PROGRAM prg_Call_Recipe_Slow
VAR
	i							: INT;
	bFirstScan					: BOOL:= TRUE;
	ton_RecipeReady				: TON;
	
	
	eRecipeName: E_Recipe_Name;

	r_trigAxisPoints_Loaded: R_TRIG;
	ton_WriteLoaded_Points: TON;
	r_trigRecipe3_loaded: R_TRIG;

	bAllRecipesLoaded: BOOL;
	iRecipeSwitchFrameVar: INT;
	bLoadDefForAll: BOOL;
	
	tPath: STRING(80);
END_VAR

act_Set_StoragePath_For_All();
//act_LoadDeafult();

ton_RecipeReady(PT:=T#1S, IN:=GVL_Recipe.stRecipe[1].bInit AND bFirstScan);
IF ton_RecipeReady.Q THEN;
	bFirstScan:=FALSE;
	bLoadDefForAll:=TRUE;
END_IF




(********************  Other Instances Recipes******************************) // 
FOR eRecipeName:=1 TO E_Recipe_Name.R_Piston_Settings DO	
	fbRecipe[eRecipeName](pstRecipe:=ADR(GVL_Recipe.stRecipe[eRecipeName]), 
			bMemoRecipeUpdated:=, 
			sRecipeDef:=TO_STRING(eRecipeName),
			bLoadDefault:=ar_RecipesLoadDefault[eRecipeName],
			bHMI_FrameActive:=iRecipeSwitchFrameVar=eRecipeName-1,//changed
			sRecipesStoragePath:=ar_RecipesStoragePath[eRecipeName]);
END_FOR
(*			
IF (*fbRecipe_1.bMemoRecipeUpdated AND*) 
fbRecipe_2.bMemoRecipeUpdated 
AND fbRecipe_3.bMemoRecipeUpdated 
AND fbRecipe_4.bMemoRecipeUpdated 
AND fbRecipe_5.bMemoRecipeUpdated 
THEN;
	bAllRecipesLoaded:=TRUE;
ELSE;
	bAllRecipesLoaded:=FALSE;
END_IF
*)

ACTION act_LoadDeafult:
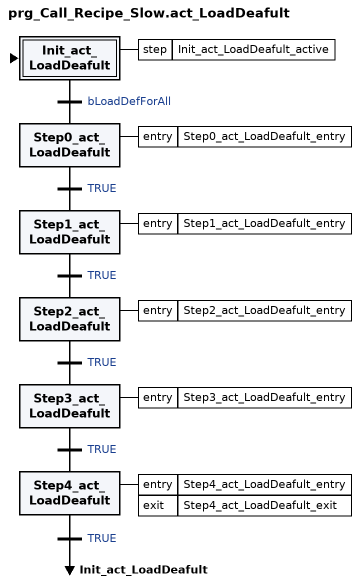
INITIAL_STEP Init_act_LoadDeafult:
    Init_act_LoadDeafult_active(N);  // step action
END_STEP
TRANSITION FROM Init_act_LoadDeafult TO Step0_act_LoadDeafult
    := bLoadDefForAll;
END_TRANSITION
STEP Step0_act_LoadDeafult:  // min time T#2s
    Step0_act_LoadDeafult_entry(P1);  // entry action
END_STEP
TRANSITION FROM Step0_act_LoadDeafult TO Step1_act_LoadDeafult
    := TRUE;
END_TRANSITION
STEP Step1_act_LoadDeafult:  // min time T#2s
    Step1_act_LoadDeafult_entry(P1);  // entry action
END_STEP
TRANSITION FROM Step1_act_LoadDeafult TO Step2_act_LoadDeafult
    := TRUE;
END_TRANSITION
STEP Step2_act_LoadDeafult:  // min time T#2s
    Step2_act_LoadDeafult_entry(P1);  // entry action
END_STEP
TRANSITION FROM Step2_act_LoadDeafult TO Step3_act_LoadDeafult
    := TRUE;
END_TRANSITION
STEP Step3_act_LoadDeafult:  // min time T#2s
    Step3_act_LoadDeafult_entry(P1);  // entry action
END_STEP
TRANSITION FROM Step3_act_LoadDeafult TO Step4_act_LoadDeafult
    := TRUE;
END_TRANSITION
STEP Step4_act_LoadDeafult:  // min time T#2s
    Step4_act_LoadDeafult_entry(P1);  // entry action
    Step4_act_LoadDeafult_exit(P0);  // exit action
END_STEP
TRANSITION FROM Step4_act_LoadDeafult TO Init_act_LoadDeafult
    := TRUE;
END_TRANSITION
END_ACTION

ACTION act_Set_StoragePath_For_All:
FOR eRecipeName:=1 TO E_Recipe_Name.R_Piston_Settings DO;
	GVL_Recipe.ar_RecipesStoragePath_Folder[eRecipeName]:=TO_STRING(eRecipeName);
	tPath:='';
	tPath:=CONCAT(tPath,GVL_Recipe.ar_RecipesStoragePath_Root[GVL_Recipe.eRecipeRootFolder]);
	tPath:=CONCAT(tPath,'\');
	tPath:=CONCAT(tPath,TO_STRING(eRecipeName));
	tPath:=CONCAT(tPath,'\');
	GVL_Recipe.ar_RecipesStoragePath[eRecipeName]:=tPath;
(*
	GVL_Recipe.ar_RecipesStoragePath[eRecipeName]:=
			CONCAT(	GVL_Recipe.ar_RecipesStoragePath_Root[GVL_Recipe.eRecipeRootFolder],'\'); 
	GVL_Recipe.ar_RecipesStoragePath[eRecipeName]:=		
			CONCAT(	GVL_Recipe.ar_RecipesStoragePath[eRecipeName],TO_STRING(eRecipeName));
	GVL_Recipe.ar_RecipesStoragePath[eRecipeName]:=		
			CONCAT(	GVL_Recipe.ar_RecipesStoragePath[eRecipeName],'1');				
	GVL_Recipe.ar_RecipesStoragePath[eRecipeName]:=		
			CONCAT(	GVL_Recipe.ar_RecipesStoragePath[eRecipeName],'\');		
*)	
END_FOR
END_ACTION

ACTION Init_act_LoadDeafult_active:
GVL_Recipe.ar_RecipesLoadDefault[1]:=FALSE;
GVL_Recipe.ar_RecipesLoadDefault[2]:=FALSE;
GVL_Recipe.ar_RecipesLoadDefault[3]:=FALSE;
GVL_Recipe.ar_RecipesLoadDefault[4]:=FALSE;
GVL_Recipe.ar_RecipesLoadDefault[5]:=FALSE;
END_ACTION

ACTION Step0_act_LoadDeafult_entry:
GVL_Recipe.ar_RecipesLoadDefault[1]:=TRUE;
END_ACTION

ACTION Step1_act_LoadDeafult_entry:
GVL_Recipe.ar_RecipesLoadDefault[2]:=TRUE;
END_ACTION

ACTION Step2_act_LoadDeafult_entry:
GVL_Recipe.ar_RecipesLoadDefault[3]:=TRUE;
END_ACTION

ACTION Step3_act_LoadDeafult_entry:
GVL_Recipe.ar_RecipesLoadDefault[4]:=TRUE;
END_ACTION

ACTION Step4_act_LoadDeafult_entry:
GVL_Recipe.ar_RecipesLoadDefault[5]:=TRUE;
END_ACTION

ACTION Step4_act_LoadDeafult_exit:
bLoadDefForAll:=FALSE;
END_ACTION

END_PROGRAM

(* stored: Version 1.1.0.1, ProductVersion 3.1.4024.12
   POU prg_Call_Recipe_Slow: Id {e80a20ed-0f91-4c74-97d3-601d773194b4}, SpecialFunc None
   Action act_LoadDeafult: Id {32d5d9ca-af5e-4d19-8254-21cc7ec9acc6}
   Action act_Set_StoragePath_For_All: Id {ab44a9a9-b46c-4897-9f85-ed22925f62ec}
   Action Init_act_LoadDeafult_active: Id {e98caf01-4c69-4303-89b4-90b4679ef1f1}
   Action Step0_act_LoadDeafult_entry: Id {a5f36d79-5c32-44ba-b9dd-e2608833fb06}
   Action Step1_act_LoadDeafult_entry: Id {d7b6e2b4-25f3-4edf-ab1a-39cc1b78fcee}
   Action Step2_act_LoadDeafult_entry: Id {0ccea3ab-e696-421c-a037-391cdca6f49f}
   Action Step3_act_LoadDeafult_entry: Id {7f0bfc77-ad46-445e-b708-4a43616e805b}
   Action Step4_act_LoadDeafult_entry: Id {043db243-9554-4cc2-887e-62028a95ea50}
   Action Step4_act_LoadDeafult_exit: Id {cb68376b-3480-475c-a045-96ddefa465d6} *)
